// Generated by voz_llm_plc_agent
// Target: Siemens TIA Portal V18 - SCL external source
// Review and compile before any download to physical hardware.

FUNCTION_BLOCK "PLC_PRG"
{ S7_Optimized_Access := 'TRUE' }
VERSION : 0.1
VAR_INPUT
   I_Emergency : Bool := FALSE;
   I_Start : Bool := FALSE;
END_VAR
VAR_OUTPUT
   Q_Motor_Enable : Bool := FALSE;
END_VAR
BEGIN
(* Arranque subordinado a la emergencia *)
#Q_Motor_Enable := #I_Start AND NOT #I_Emergency;
(* Prioridad absoluta del paro de emergencia *)
IF #I_Emergency THEN
    #Q_Motor_Enable := FALSE;
END_IF;
END_FUNCTION_BLOCK

DATA_BLOCK "DB_PLC_PRG"
{ S7_Optimized_Access := 'TRUE' }
VERSION : 0.1
NON_RETAIN
"PLC_PRG"
BEGIN
END_DATA_BLOCK

ORGANIZATION_BLOCK "Main"
{ S7_Optimized_Access := 'TRUE' }
VERSION : 0.1
BEGIN
   "DB_PLC_PRG"(
      I_Emergency := "I_Emergency",
      Q_Motor_Enable => "Q_Motor_Enable",
      I_Start := "I_Start"
   );
END_ORGANIZATION_BLOCK
